// TIA Portal V20 export
// export: Created 2026-10-12T05:00:30.1846246Z, ExportSetting WithDefaults, DisplayName Totally Integrated Automation Portal, DisplayVersion V20, DisplayName TIA Portal Openness, DisplayVersion V20, DisplayName TIA Portal Teamcenter Gateway, DisplayVersion V20, DisplayName TIA Portal Version Control Interface, DisplayVersion V20, DisplayName SINAMICS Startdrive Advanced, DisplayVersion V20 SP1 Update 2, DisplayName SINAMICS Startdrive G110M, G120, G120C, G120D, G120P, G115D, DisplayVersion V20 SP1 Update 2, DisplayName SINAMICS Startdrive G130, G150, S120, S150, SINAMICS MV, G220, S200, S210, DisplayVersion V20 SP1 Update 2, DisplayName STEP 7 Professional, DisplayVersion V20, DisplayName STEP 7 Safety, DisplayVersion V20, DisplayName WinCC Basic/Comfort/Advanced, DisplayVersion V20, DisplayName WinCC Professional, DisplayVersion V20, DisplayName WinCC Unified, DisplayVersion V20
FUNCTION "FRK_SetShape" : Bool   // FC112, SCL
{ S7_Optimized_Access := 'TRUE' }
VERSION : 0.1
// stored: AutoNumber true, IsIECCheckEnabled false, SetENOAutomatically false, UDAEnableTagReadback false
   VAR_INPUT
      RootIndex : Int;
      RootIdentity : String;
   END_VAR
   VAR_TEMP
      Index : Int;
      Other : Int;
      ModelIndex : Int;
      KnownModel : Bool;
   END_VAR
BEGIN

   #FRK_SetShape := FALSE;
   IF NOT "FRK_SetRuntime".Work[#RootIndex].Payload.Info.Used OR "FRK_SetRuntime".Work[#RootIndex].Payload.Info.RootIdentity <> #RootIdentity
       OR "FRK_SetRuntime".Work[#RootIndex].Payload.Info.SetSchema <> 1 OR "FRK_SetRuntime".Work[#RootIndex].Payload.Info.ConfigRev = 0
       OR LEN("FRK_SetRuntime".Work[#RootIndex].Payload.Info.SetName) = 0
       OR "FRK_SetRuntime".Work[#RootIndex].Payload.Info.RecordCount < 1 OR "FRK_SetRuntime".Work[#RootIndex].Payload.Info.RecordCount > 24 THEN
       RETURN;
   END_IF;
   IF "FRK_SetRuntime".Work[#RootIndex].Payload.Info.Kind = 0 THEN
       #KnownModel := FALSE;
       FOR #ModelIndex := 1 TO 2 DO
           IF "FRK_SetRuntime".Work[#RootIndex].Payload.Info.ModelCode = "FRK_ConfigModelCode"(RootIndex := #RootIndex, ModelIndex := INT_TO_UDINT(#ModelIndex)) THEN
               #KnownModel := TRUE;
           END_IF;
       END_FOR;
       IF NOT #KnownModel THEN
           RETURN;
       END_IF;
   ELSIF "FRK_SetRuntime".Work[#RootIndex].Payload.Info.Kind <> 1 OR "FRK_SetRuntime".Work[#RootIndex].Payload.Info.ModelCode <> '' THEN
       RETURN;
   END_IF;
   FOR #Index := 1 TO "FRK_SetRuntime".Work[#RootIndex].Payload.Info.RecordCount DO
       "FRK_SetRuntime".Work[#RootIndex].RejectScope := "FRK_SetRuntime".Work[#RootIndex].Payload.Records[#Index].Scope;
       "FRK_SetRuntime".Work[#RootIndex].RejectKey := "FRK_SetRuntime".Work[#RootIndex].Payload.Records[#Index].WriteKey;
       IF "FRK_SetRuntime".Work[#RootIndex].Payload.Records[#Index].Kind <> "FRK_SetRuntime".Work[#RootIndex].Payload.Info.Kind THEN
           RETURN;
       END_IF;
       FOR #Other := 1 TO #Index - 1 DO
           IF "FRK_SetRuntime".Work[#RootIndex].Payload.Records[#Other].Scope = "FRK_SetRuntime".Work[#RootIndex].Payload.Records[#Index].Scope
               AND "FRK_SetRuntime".Work[#RootIndex].Payload.Records[#Other].WriteKey = "FRK_SetRuntime".Work[#RootIndex].Payload.Records[#Index].WriteKey THEN
               RETURN;
           END_IF;
       END_FOR;
   END_FOR;
   #FRK_SetShape := TRUE;
END_FUNCTION
